(* PLC project failsafe_motor_latch, Unknown Lessons in Electric Circuits transcription 1 *)
(* stored: creationDateTime 2026-09-02T12:00:00 *)

PROGRAM main
  VAR
    START : BOOL;
    THERMAL_OVERLOAD_NC : BOOL;
    STOP_NC : BOOL;
    MOTOR_RUN : BOOL;
  END_VAR

(* LD diagram, written out as Structured Text *)
MOTOR_RUN := (START OR MOTOR_RUN) AND THERMAL_OVERLOAD_NC AND STOP_NC;
END_PROGRAM

CONFIGURATION Config0
  RESOURCE Res0 ON PLC
    TASK tcyclic(INTERVAL := T#10ms, PRIORITY := 0);
    PROGRAM inst0 WITH tcyclic : main;
  END_RESOURCE
END_CONFIGURATION
